// TIA Portal V19 export
FUNCTION_BLOCK "SKIDS"   // FB18, LAD
{ S7_Optimized_Access := 'TRUE' }
// stored: MemoryReserve 100, SetENOAutomatically false
   VAR
      CHILLED_SKIDS_Instance { S7_SetPoint := 'True'} : "SKIDS_LOGIC";
      START_Instance { S7_SetPoint := 'True'} : "START";
      START_Instance_COLD_SKIDS { S7_SetPoint := 'True'} : "START";
      CS_SKIDS_Instance_1 { S7_SetPoint := 'True'} : "SKIDS_LOGIC";
      START_Instance_UCH { S7_SetPoint := 'True'} : "START";
      ULTRACHILLED_SKIDS_Instance { S7_SetPoint := 'True'} : "SKIDS_LOGIC";
      ULTRACHILLED_SKIDS_Instance_1 { S7_SetPoint := 'True'} : "ULTRACHILLED_SKIDS";
      HOT_SKIDS_InstancE { S7_SetPoint := 'True'} : "SKIDS_LOGIC";
      HOT_SKIDS_Instance_1 { S7_SetPoint := 'True'} : "HOT_SKIDS";
      START_Instance_HOT_SKIDS { S7_SetPoint := 'True'} : "START";
   END_VAR
BEGIN

REGION Network 1: CHILLED SKIDS START
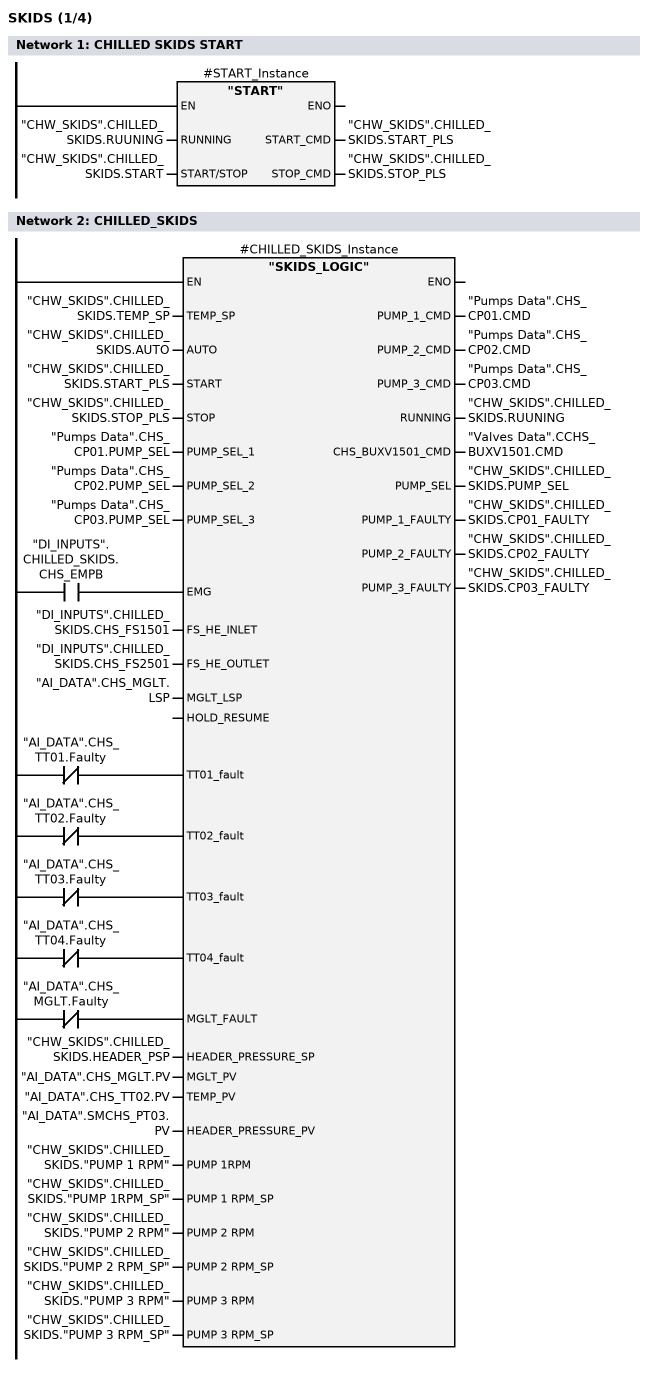
   RUNG wire#powerrail
      #START_Instance(RUNNING := "CHW_SKIDS".CHILLED_SKIDS.RUUNING, "START/STOP" := "CHW_SKIDS".CHILLED_SKIDS.START, START_CMD => "CHW_SKIDS".CHILLED_SKIDS.START_PLS, STOP_CMD => "CHW_SKIDS".CHILLED_SKIDS.STOP_PLS)
   END_RUNG
   // the same network as SCL:
   #START_Instance(RUNNING := "CHW_SKIDS".CHILLED_SKIDS.RUUNING,   // "START"
                   "START/STOP" := "CHW_SKIDS".CHILLED_SKIDS.START,
                   START_CMD => "CHW_SKIDS".CHILLED_SKIDS.START_PLS,
                   STOP_CMD => "CHW_SKIDS".CHILLED_SKIDS.STOP_PLS);
END_REGION

REGION Network 2: CHILLED_SKIDS
   RUNG wire#powerrail
      #CHILLED_SKIDS_Instance(EMG := wire#w1, TT01_fault := wire#w2, TT02_fault := wire#w3, TT03_fault := wire#w4, TT04_fault := wire#w5, MGLT_FAULT := wire#w6, TEMP_SP := "CHW_SKIDS".CHILLED_SKIDS.TEMP_SP, AUTO := "CHW_SKIDS".CHILLED_SKIDS.AUTO, START := "CHW_SKIDS".CHILLED_SKIDS.START_PLS, STOP := "CHW_SKIDS".CHILLED_SKIDS.STOP_PLS, PUMP_SEL_1 := "Pumps Data".CHS_CP01.PUMP_SEL, PUMP_SEL_2 := "Pumps Data".CHS_CP02.PUMP_SEL, PUMP_SEL_3 := "Pumps Data".CHS_CP03.PUMP_SEL, FS_HE_INLET := "DI_INPUTS".CHILLED_SKIDS.CHS_FS1501, FS_HE_OUTLET := "DI_INPUTS".CHILLED_SKIDS.CHS_FS2501, MGLT_LSP := "AI_DATA".CHS_MGLT.LSP, HOLD_RESUME :=, HEADER_PRESSURE_SP := "CHW_SKIDS".CHILLED_SKIDS.HEADER_PSP, MGLT_PV := "AI_DATA".CHS_MGLT.PV, TEMP_PV := "AI_DATA".CHS_TT02.PV, HEADER_PRESSURE_PV := "AI_DATA".SMCHS_PT03.PV, "PUMP 1RPM" := "CHW_SKIDS".CHILLED_SKIDS."PUMP 1 RPM", "PUMP 1 RPM_SP" := "CHW_SKIDS".CHILLED_SKIDS."PUMP 1RPM_SP", "PUMP 2 RPM" := "CHW_SKIDS".CHILLED_SKIDS."PUMP 2 RPM", "PUMP 2 RPM_SP" := "CHW_SKIDS".CHILLED_SKIDS."PUMP 2 RPM_SP", "PUMP 3 RPM" := "CHW_SKIDS".CHILLED_SKIDS."PUMP 3 RPM", "PUMP 3 RPM_SP" := "CHW_SKIDS".CHILLED_SKIDS."PUMP 3 RPM_SP", PUMP_1_CMD => "Pumps Data".CHS_CP01.CMD, PUMP_2_CMD => "Pumps Data".CHS_CP02.CMD, PUMP_3_CMD => "Pumps Data".CHS_CP03.CMD, RUNNING => "CHW_SKIDS".CHILLED_SKIDS.RUUNING, CHS_BUXV1501_CMD => "Valves Data".CCHS_BUXV1501.CMD, PUMP_SEL => "CHW_SKIDS".CHILLED_SKIDS.PUMP_SEL, PUMP_1_FAULTY => "CHW_SKIDS".CHILLED_SKIDS.CP01_FAULTY, PUMP_2_FAULTY => "CHW_SKIDS".CHILLED_SKIDS.CP02_FAULTY, PUMP_3_FAULTY => "CHW_SKIDS".CHILLED_SKIDS.CP03_FAULTY)
   END_RUNG
   RUNG wire#powerrail
      Contact( "DI_INPUTS".CHILLED_SKIDS.CHS_EMPB )
   END_RUNG wire#w1
   RUNG wire#powerrail
      I_Contact( "AI_DATA".CHS_TT01.Faulty )
   END_RUNG wire#w2
   RUNG wire#powerrail
      I_Contact( "AI_DATA".CHS_TT02.Faulty )
   END_RUNG wire#w3
   RUNG wire#powerrail
      I_Contact( "AI_DATA".CHS_TT03.Faulty )
   END_RUNG wire#w4
   RUNG wire#powerrail
      I_Contact( "AI_DATA".CHS_TT04.Faulty )
   END_RUNG wire#w5
   RUNG wire#powerrail
      I_Contact( "AI_DATA".CHS_MGLT.Faulty )
   END_RUNG wire#w6
   // the same network as SCL:
   #CHILLED_SKIDS_Instance(TEMP_SP := "CHW_SKIDS".CHILLED_SKIDS.TEMP_SP,   // "SKIDS_LOGIC"
                           AUTO := "CHW_SKIDS".CHILLED_SKIDS.AUTO,
                           START := "CHW_SKIDS".CHILLED_SKIDS.START_PLS,
                           STOP := "CHW_SKIDS".CHILLED_SKIDS.STOP_PLS,
                           PUMP_SEL_1 := "Pumps Data".CHS_CP01.PUMP_SEL,
                           PUMP_SEL_2 := "Pumps Data".CHS_CP02.PUMP_SEL,
                           PUMP_SEL_3 := "Pumps Data".CHS_CP03.PUMP_SEL,
                           EMG := "DI_INPUTS".CHILLED_SKIDS.CHS_EMPB,
                           FS_HE_INLET := "DI_INPUTS".CHILLED_SKIDS.CHS_FS1501,
                           FS_HE_OUTLET := "DI_INPUTS".CHILLED_SKIDS.CHS_FS2501,
                           MGLT_LSP := "AI_DATA".CHS_MGLT.LSP,
                           TT01_fault := NOT "AI_DATA".CHS_TT01.Faulty,
                           TT02_fault := NOT "AI_DATA".CHS_TT02.Faulty,
                           TT03_fault := NOT "AI_DATA".CHS_TT03.Faulty,
                           TT04_fault := NOT "AI_DATA".CHS_TT04.Faulty,
                           MGLT_FAULT := NOT "AI_DATA".CHS_MGLT.Faulty,
                           HEADER_PRESSURE_SP := "CHW_SKIDS".CHILLED_SKIDS.HEADER_PSP,
                           MGLT_PV := "AI_DATA".CHS_MGLT.PV,
                           TEMP_PV := "AI_DATA".CHS_TT02.PV,
                           HEADER_PRESSURE_PV := "AI_DATA".SMCHS_PT03.PV,
                           "PUMP 1RPM" := "CHW_SKIDS".CHILLED_SKIDS."PUMP 1 RPM",
                           "PUMP 1 RPM_SP" := "CHW_SKIDS".CHILLED_SKIDS."PUMP 1RPM_SP",
                           "PUMP 2 RPM" := "CHW_SKIDS".CHILLED_SKIDS."PUMP 2 RPM",
                           "PUMP 2 RPM_SP" := "CHW_SKIDS".CHILLED_SKIDS."PUMP 2 RPM_SP",
                           "PUMP 3 RPM" := "CHW_SKIDS".CHILLED_SKIDS."PUMP 3 RPM",
                           "PUMP 3 RPM_SP" := "CHW_SKIDS".CHILLED_SKIDS."PUMP 3 RPM_SP",
                           PUMP_1_CMD => "Pumps Data".CHS_CP01.CMD,
                           PUMP_2_CMD => "Pumps Data".CHS_CP02.CMD,
                           PUMP_3_CMD => "Pumps Data".CHS_CP03.CMD,
                           RUNNING => "CHW_SKIDS".CHILLED_SKIDS.RUUNING,
                           CHS_BUXV1501_CMD => "Valves Data".CCHS_BUXV1501.CMD,
                           PUMP_SEL => "CHW_SKIDS".CHILLED_SKIDS.PUMP_SEL,
                           PUMP_1_FAULTY => "CHW_SKIDS".CHILLED_SKIDS.CP01_FAULTY,
                           PUMP_2_FAULTY => "CHW_SKIDS".CHILLED_SKIDS.CP02_FAULTY,
                           PUMP_3_FAULTY => "CHW_SKIDS".CHILLED_SKIDS.CP03_FAULTY);
END_REGION

REGION Network 3: COLD SKIDS START
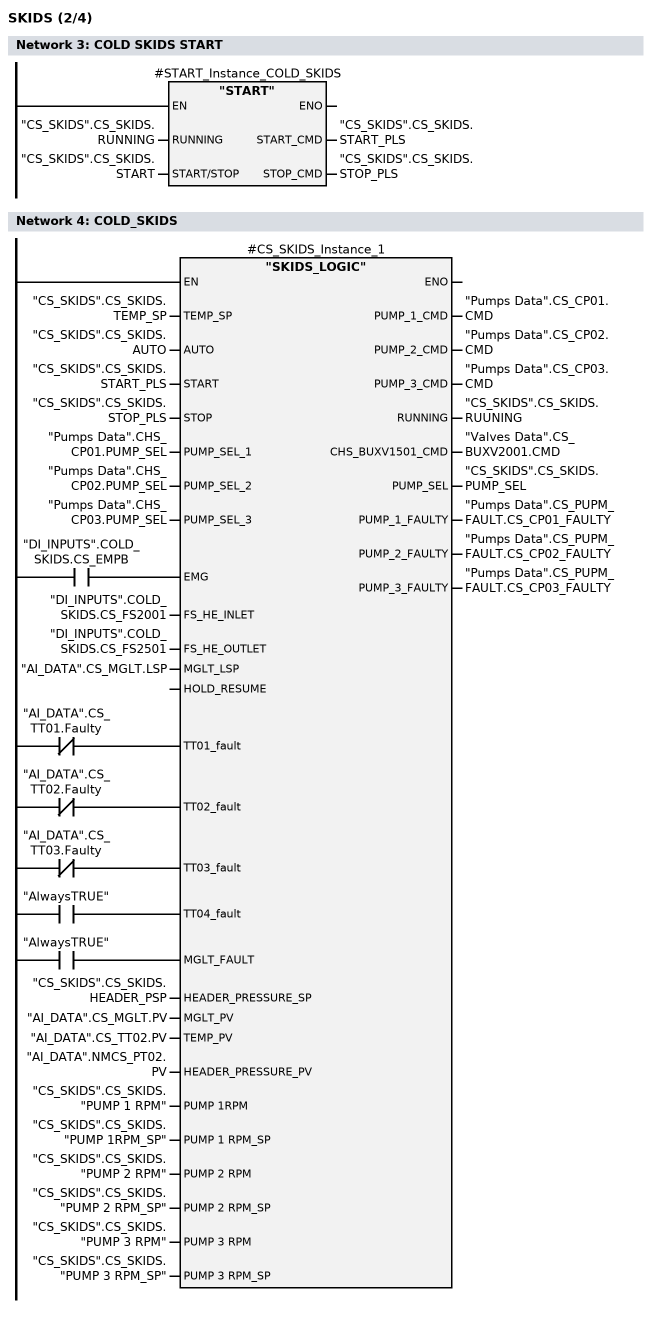
   RUNG wire#powerrail
      #START_Instance_COLD_SKIDS(RUNNING := "CS_SKIDS".CS_SKIDS.RUNNING, "START/STOP" := "CS_SKIDS".CS_SKIDS.START, START_CMD => "CS_SKIDS".CS_SKIDS.START_PLS, STOP_CMD => "CS_SKIDS".CS_SKIDS.STOP_PLS)
   END_RUNG
   // the same network as SCL:
   #START_Instance_COLD_SKIDS(RUNNING := "CS_SKIDS".CS_SKIDS.RUNNING,   // "START"
                           "START/STOP" := "CS_SKIDS".CS_SKIDS.START,
                           START_CMD => "CS_SKIDS".CS_SKIDS.START_PLS,
                           STOP_CMD => "CS_SKIDS".CS_SKIDS.STOP_PLS);
END_REGION

REGION Network 4: COLD_SKIDS
   RUNG wire#powerrail
      #CS_SKIDS_Instance_1(EMG := wire#w1, TT01_fault := wire#w2, TT02_fault := wire#w3, TT03_fault := wire#w4, TT04_fault := wire#w5, MGLT_FAULT := wire#w6, TEMP_SP := "CS_SKIDS".CS_SKIDS.TEMP_SP, AUTO := "CS_SKIDS".CS_SKIDS.AUTO, START := "CS_SKIDS".CS_SKIDS.START_PLS, STOP := "CS_SKIDS".CS_SKIDS.STOP_PLS, PUMP_SEL_1 := "Pumps Data".CHS_CP01.PUMP_SEL, PUMP_SEL_2 := "Pumps Data".CHS_CP02.PUMP_SEL, PUMP_SEL_3 := "Pumps Data".CHS_CP03.PUMP_SEL, FS_HE_INLET := "DI_INPUTS".COLD_SKIDS.CS_FS2001, FS_HE_OUTLET := "DI_INPUTS".COLD_SKIDS.CS_FS2501, MGLT_LSP := "AI_DATA".CS_MGLT.LSP, HOLD_RESUME :=, HEADER_PRESSURE_SP := "CS_SKIDS".CS_SKIDS.HEADER_PSP, MGLT_PV := "AI_DATA".CS_MGLT.PV, TEMP_PV := "AI_DATA".CS_TT02.PV, HEADER_PRESSURE_PV := "AI_DATA".NMCS_PT02.PV, "PUMP 1RPM" := "CS_SKIDS".CS_SKIDS."PUMP 1 RPM", "PUMP 1 RPM_SP" := "CS_SKIDS".CS_SKIDS."PUMP 1RPM_SP", "PUMP 2 RPM" := "CS_SKIDS".CS_SKIDS."PUMP 2 RPM", "PUMP 2 RPM_SP" := "CS_SKIDS".CS_SKIDS."PUMP 2 RPM_SP", "PUMP 3 RPM" := "CS_SKIDS".CS_SKIDS."PUMP 3 RPM", "PUMP 3 RPM_SP" := "CS_SKIDS".CS_SKIDS."PUMP 3 RPM_SP", PUMP_1_CMD => "Pumps Data".CS_CP01.CMD, PUMP_2_CMD => "Pumps Data".CS_CP02.CMD, PUMP_3_CMD => "Pumps Data".CS_CP03.CMD, RUNNING => "CS_SKIDS".CS_SKIDS.RUUNING, CHS_BUXV1501_CMD => "Valves Data".CS_BUXV2001.CMD, PUMP_SEL => "CS_SKIDS".CS_SKIDS.PUMP_SEL, PUMP_1_FAULTY => "Pumps Data".CS_PUPM_FAULT.CS_CP01_FAULTY, PUMP_2_FAULTY => "Pumps Data".CS_PUPM_FAULT.CS_CP02_FAULTY, PUMP_3_FAULTY => "Pumps Data".CS_PUPM_FAULT.CS_CP03_FAULTY)
   END_RUNG
   RUNG wire#powerrail
      Contact( "DI_INPUTS".COLD_SKIDS.CS_EMPB )
   END_RUNG wire#w1
   RUNG wire#powerrail
      I_Contact( "AI_DATA".CS_TT01.Faulty )
   END_RUNG wire#w2
   RUNG wire#powerrail
      I_Contact( "AI_DATA".CS_TT02.Faulty )
   END_RUNG wire#w3
   RUNG wire#powerrail
      I_Contact( "AI_DATA".CS_TT03.Faulty )
   END_RUNG wire#w4
   RUNG wire#powerrail
      Contact( "AlwaysTRUE" )
   END_RUNG wire#w5
   RUNG wire#powerrail
      Contact( "AlwaysTRUE" )
   END_RUNG wire#w6
   // the same network as SCL:
   #CS_SKIDS_Instance_1(TEMP_SP := "CS_SKIDS".CS_SKIDS.TEMP_SP,   // "SKIDS_LOGIC"
                        AUTO := "CS_SKIDS".CS_SKIDS.AUTO,
                        START := "CS_SKIDS".CS_SKIDS.START_PLS,
                        STOP := "CS_SKIDS".CS_SKIDS.STOP_PLS,
                        PUMP_SEL_1 := "Pumps Data".CHS_CP01.PUMP_SEL,
                        PUMP_SEL_2 := "Pumps Data".CHS_CP02.PUMP_SEL,
                        PUMP_SEL_3 := "Pumps Data".CHS_CP03.PUMP_SEL,
                        EMG := "DI_INPUTS".COLD_SKIDS.CS_EMPB,
                        FS_HE_INLET := "DI_INPUTS".COLD_SKIDS.CS_FS2001,
                        FS_HE_OUTLET := "DI_INPUTS".COLD_SKIDS.CS_FS2501,
                        MGLT_LSP := "AI_DATA".CS_MGLT.LSP,
                        TT01_fault := NOT "AI_DATA".CS_TT01.Faulty,
                        TT02_fault := NOT "AI_DATA".CS_TT02.Faulty,
                        TT03_fault := NOT "AI_DATA".CS_TT03.Faulty,
                        TT04_fault := "AlwaysTRUE",
                        MGLT_FAULT := "AlwaysTRUE",
                        HEADER_PRESSURE_SP := "CS_SKIDS".CS_SKIDS.HEADER_PSP,
                        MGLT_PV := "AI_DATA".CS_MGLT.PV,
                        TEMP_PV := "AI_DATA".CS_TT02.PV,
                        HEADER_PRESSURE_PV := "AI_DATA".NMCS_PT02.PV,
                        "PUMP 1RPM" := "CS_SKIDS".CS_SKIDS."PUMP 1 RPM",
                        "PUMP 1 RPM_SP" := "CS_SKIDS".CS_SKIDS."PUMP 1RPM_SP",
                        "PUMP 2 RPM" := "CS_SKIDS".CS_SKIDS."PUMP 2 RPM",
                        "PUMP 2 RPM_SP" := "CS_SKIDS".CS_SKIDS."PUMP 2 RPM_SP",
                        "PUMP 3 RPM" := "CS_SKIDS".CS_SKIDS."PUMP 3 RPM",
                        "PUMP 3 RPM_SP" := "CS_SKIDS".CS_SKIDS."PUMP 3 RPM_SP",
                        PUMP_1_CMD => "Pumps Data".CS_CP01.CMD,
                        PUMP_2_CMD => "Pumps Data".CS_CP02.CMD,
                        PUMP_3_CMD => "Pumps Data".CS_CP03.CMD,
                        RUNNING => "CS_SKIDS".CS_SKIDS.RUUNING,
                        CHS_BUXV1501_CMD => "Valves Data".CS_BUXV2001.CMD,
                        PUMP_SEL => "CS_SKIDS".CS_SKIDS.PUMP_SEL,
                        PUMP_1_FAULTY => "Pumps Data".CS_PUPM_FAULT.CS_CP01_FAULTY,
                        PUMP_2_FAULTY => "Pumps Data".CS_PUPM_FAULT.CS_CP02_FAULTY,
                        PUMP_3_FAULTY => "Pumps Data".CS_PUPM_FAULT.CS_CP03_FAULTY);
END_REGION

REGION Network 5: ULTRACHILLED SKIDS START
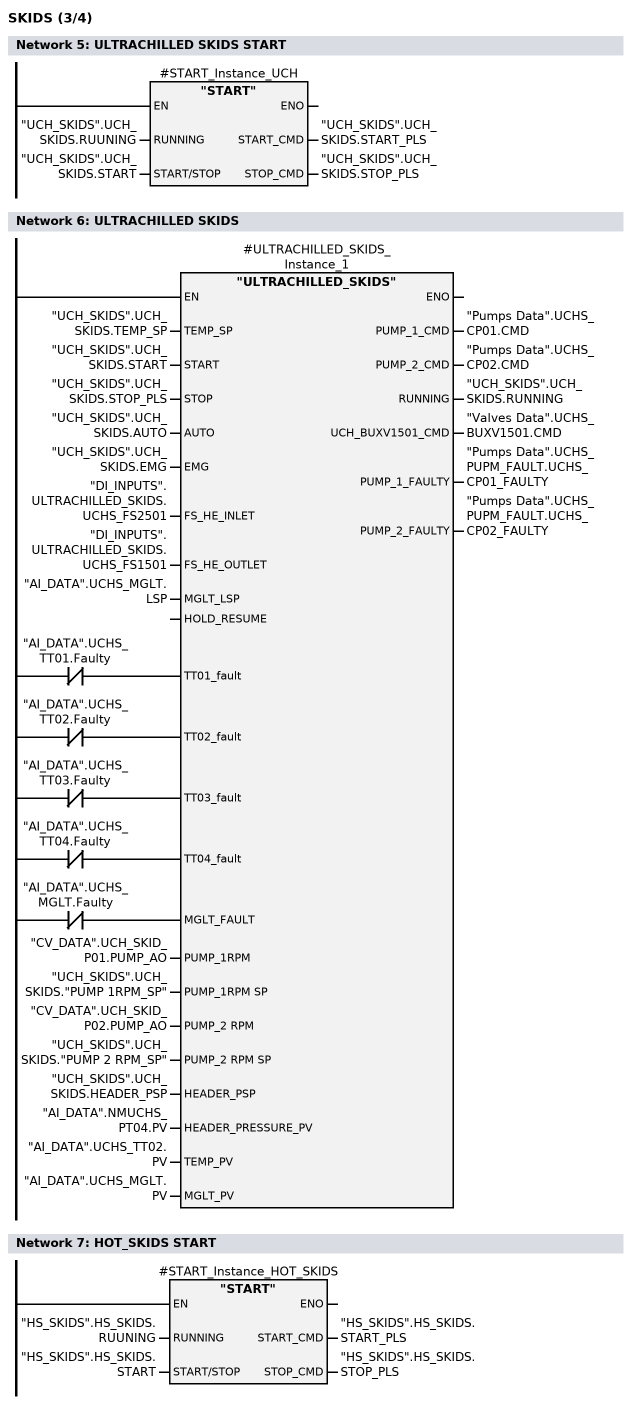
   RUNG wire#powerrail
      #START_Instance_UCH(RUNNING := "UCH_SKIDS".UCH_SKIDS.RUUNING, "START/STOP" := "UCH_SKIDS".UCH_SKIDS.START, START_CMD => "UCH_SKIDS".UCH_SKIDS.START_PLS, STOP_CMD => "UCH_SKIDS".UCH_SKIDS.STOP_PLS)
   END_RUNG
   // the same network as SCL:
   #START_Instance_UCH(RUNNING := "UCH_SKIDS".UCH_SKIDS.RUUNING,   // "START"
                       "START/STOP" := "UCH_SKIDS".UCH_SKIDS.START,
                       START_CMD => "UCH_SKIDS".UCH_SKIDS.START_PLS,
                       STOP_CMD => "UCH_SKIDS".UCH_SKIDS.STOP_PLS);
END_REGION

REGION Network 6: ULTRACHILLED SKIDS
   RUNG wire#powerrail
      #ULTRACHILLED_SKIDS_Instance_1(TT01_fault := wire#w1, TT02_fault := wire#w2, TT03_fault := wire#w3, TT04_fault := wire#w4, MGLT_FAULT := wire#w5, TEMP_SP := "UCH_SKIDS".UCH_SKIDS.TEMP_SP, START := "UCH_SKIDS".UCH_SKIDS.START, STOP := "UCH_SKIDS".UCH_SKIDS.STOP_PLS, AUTO := "UCH_SKIDS".UCH_SKIDS.AUTO, EMG := "UCH_SKIDS".UCH_SKIDS.EMG, FS_HE_INLET := "DI_INPUTS".ULTRACHILLED_SKIDS.UCHS_FS2501, FS_HE_OUTLET := "DI_INPUTS".ULTRACHILLED_SKIDS.UCHS_FS1501, MGLT_LSP := "AI_DATA".UCHS_MGLT.LSP, HOLD_RESUME :=, PUMP_1RPM := "CV_DATA".UCH_SKID_P01.PUMP_AO, "PUMP_1RPM SP" := "UCH_SKIDS".UCH_SKIDS."PUMP 1RPM_SP", "PUMP_2 RPM" := "CV_DATA".UCH_SKID_P02.PUMP_AO, "PUMP_2 RPM SP" := "UCH_SKIDS".UCH_SKIDS."PUMP 2 RPM_SP", HEADER_PSP := "UCH_SKIDS".UCH_SKIDS.HEADER_PSP, HEADER_PRESSURE_PV := "AI_DATA".NMUCHS_PT04.PV, TEMP_PV := "AI_DATA".UCHS_TT02.PV, MGLT_PV := "AI_DATA".UCHS_MGLT.PV, PUMP_1_CMD => "Pumps Data".UCHS_CP01.CMD, PUMP_2_CMD => "Pumps Data".UCHS_CP02.CMD, RUNNING => "UCH_SKIDS".UCH_SKIDS.RUNNING, UCH_BUXV1501_CMD => "Valves Data".UCHS_BUXV1501.CMD, PUMP_1_FAULTY => "Pumps Data".UCHS_PUPM_FAULT.UCHS_CP01_FAULTY, PUMP_2_FAULTY => "Pumps Data".UCHS_PUPM_FAULT.UCHS_CP02_FAULTY)
   END_RUNG
   RUNG wire#powerrail
      I_Contact( "AI_DATA".UCHS_TT01.Faulty )
   END_RUNG wire#w1
   RUNG wire#powerrail
      I_Contact( "AI_DATA".UCHS_TT02.Faulty )
   END_RUNG wire#w2
   RUNG wire#powerrail
      I_Contact( "AI_DATA".UCHS_TT03.Faulty )
   END_RUNG wire#w3
   RUNG wire#powerrail
      I_Contact( "AI_DATA".UCHS_TT04.Faulty )
   END_RUNG wire#w4
   RUNG wire#powerrail
      I_Contact( "AI_DATA".UCHS_MGLT.Faulty )
   END_RUNG wire#w5
   // the same network as SCL:
   #ULTRACHILLED_SKIDS_Instance_1(TEMP_SP := "UCH_SKIDS".UCH_SKIDS.TEMP_SP,   // "ULTRACHILLED_SKIDS"
                           START := "UCH_SKIDS".UCH_SKIDS.START,
                           STOP := "UCH_SKIDS".UCH_SKIDS.STOP_PLS,
                           AUTO := "UCH_SKIDS".UCH_SKIDS.AUTO,
                           EMG := "UCH_SKIDS".UCH_SKIDS.EMG,
                           FS_HE_INLET := "DI_INPUTS".ULTRACHILLED_SKIDS.UCHS_FS2501,
                           FS_HE_OUTLET := "DI_INPUTS".ULTRACHILLED_SKIDS.UCHS_FS1501,
                           MGLT_LSP := "AI_DATA".UCHS_MGLT.LSP,
                           TT01_fault := NOT "AI_DATA".UCHS_TT01.Faulty,
                           TT02_fault := NOT "AI_DATA".UCHS_TT02.Faulty,
                           TT03_fault := NOT "AI_DATA".UCHS_TT03.Faulty,
                           TT04_fault := NOT "AI_DATA".UCHS_TT04.Faulty,
                           MGLT_FAULT := NOT "AI_DATA".UCHS_MGLT.Faulty,
                           PUMP_1RPM := "CV_DATA".UCH_SKID_P01.PUMP_AO,
                           "PUMP_1RPM SP" := "UCH_SKIDS".UCH_SKIDS."PUMP 1RPM_SP",
                           "PUMP_2 RPM" := "CV_DATA".UCH_SKID_P02.PUMP_AO,
                           "PUMP_2 RPM SP" := "UCH_SKIDS".UCH_SKIDS."PUMP 2 RPM_SP",
                           HEADER_PSP := "UCH_SKIDS".UCH_SKIDS.HEADER_PSP,
                           HEADER_PRESSURE_PV := "AI_DATA".NMUCHS_PT04.PV,
                           TEMP_PV := "AI_DATA".UCHS_TT02.PV,
                           MGLT_PV := "AI_DATA".UCHS_MGLT.PV,
                           PUMP_1_CMD => "Pumps Data".UCHS_CP01.CMD,
                           PUMP_2_CMD => "Pumps Data".UCHS_CP02.CMD,
                           RUNNING => "UCH_SKIDS".UCH_SKIDS.RUNNING,
                           UCH_BUXV1501_CMD => "Valves Data".UCHS_BUXV1501.CMD,
                           PUMP_1_FAULTY => "Pumps Data".UCHS_PUPM_FAULT.UCHS_CP01_FAULTY,
                           PUMP_2_FAULTY => "Pumps Data".UCHS_PUPM_FAULT.UCHS_CP02_FAULTY);
END_REGION

REGION Network 7: HOT_SKIDS START
   RUNG wire#powerrail
      #START_Instance_HOT_SKIDS(RUNNING := "HS_SKIDS".HS_SKIDS.RUUNING, "START/STOP" := "HS_SKIDS".HS_SKIDS.START, START_CMD => "HS_SKIDS".HS_SKIDS.START_PLS, STOP_CMD => "HS_SKIDS".HS_SKIDS.STOP_PLS)
   END_RUNG
   // the same network as SCL:
   #START_Instance_HOT_SKIDS(RUNNING := "HS_SKIDS".HS_SKIDS.RUUNING,   // "START"
                           "START/STOP" := "HS_SKIDS".HS_SKIDS.START,
                           START_CMD => "HS_SKIDS".HS_SKIDS.START_PLS,
                           STOP_CMD => "HS_SKIDS".HS_SKIDS.STOP_PLS);
END_REGION

REGION Network 8: HOT_SKIDS
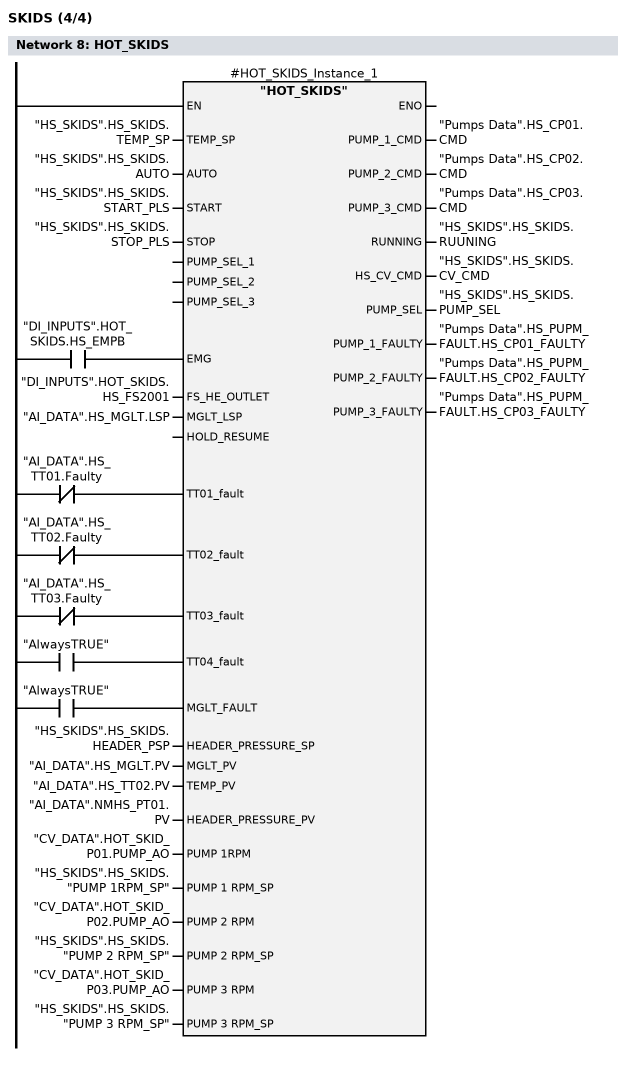
   RUNG wire#powerrail
      #HOT_SKIDS_Instance_1(EMG := wire#w1, TT01_fault := wire#w2, TT02_fault := wire#w3, TT03_fault := wire#w4, TT04_fault := wire#w5, MGLT_FAULT := wire#w6, TEMP_SP := "HS_SKIDS".HS_SKIDS.TEMP_SP, AUTO := "HS_SKIDS".HS_SKIDS.AUTO, START := "HS_SKIDS".HS_SKIDS.START_PLS, STOP := "HS_SKIDS".HS_SKIDS.STOP_PLS, PUMP_SEL_1 :=, PUMP_SEL_2 :=, PUMP_SEL_3 :=, FS_HE_OUTLET := "DI_INPUTS".HOT_SKIDS.HS_FS2001, MGLT_LSP := "AI_DATA".HS_MGLT.LSP, HOLD_RESUME :=, HEADER_PRESSURE_SP := "HS_SKIDS".HS_SKIDS.HEADER_PSP, MGLT_PV := "AI_DATA".HS_MGLT.PV, TEMP_PV := "AI_DATA".HS_TT02.PV, HEADER_PRESSURE_PV := "AI_DATA".NMHS_PT01.PV, "PUMP 1RPM" := "CV_DATA".HOT_SKID_P01.PUMP_AO, "PUMP 1 RPM_SP" := "HS_SKIDS".HS_SKIDS."PUMP 1RPM_SP", "PUMP 2 RPM" := "CV_DATA".HOT_SKID_P02.PUMP_AO, "PUMP 2 RPM_SP" := "HS_SKIDS".HS_SKIDS."PUMP 2 RPM_SP", "PUMP 3 RPM" := "CV_DATA".HOT_SKID_P03.PUMP_AO, "PUMP 3 RPM_SP" := "HS_SKIDS".HS_SKIDS."PUMP 3 RPM_SP", PUMP_1_CMD => "Pumps Data".HS_CP01.CMD, PUMP_2_CMD => "Pumps Data".HS_CP02.CMD, PUMP_3_CMD => "Pumps Data".HS_CP03.CMD, RUNNING => "HS_SKIDS".HS_SKIDS.RUUNING, HS_CV_CMD => "HS_SKIDS".HS_SKIDS.CV_CMD, PUMP_SEL => "HS_SKIDS".HS_SKIDS.PUMP_SEL, PUMP_1_FAULTY => "Pumps Data".HS_PUPM_FAULT.HS_CP01_FAULTY, PUMP_2_FAULTY => "Pumps Data".HS_PUPM_FAULT.HS_CP02_FAULTY, PUMP_3_FAULTY => "Pumps Data".HS_PUPM_FAULT.HS_CP03_FAULTY)
   END_RUNG
   RUNG wire#powerrail
      Contact( "DI_INPUTS".HOT_SKIDS.HS_EMPB )
   END_RUNG wire#w1
   RUNG wire#powerrail
      I_Contact( "AI_DATA".HS_TT01.Faulty )
   END_RUNG wire#w2
   RUNG wire#powerrail
      I_Contact( "AI_DATA".HS_TT02.Faulty )
   END_RUNG wire#w3
   RUNG wire#powerrail
      I_Contact( "AI_DATA".HS_TT03.Faulty )
   END_RUNG wire#w4
   RUNG wire#powerrail
      Contact( "AlwaysTRUE" )
   END_RUNG wire#w5
   RUNG wire#powerrail
      Contact( "AlwaysTRUE" )
   END_RUNG wire#w6
   // the same network as SCL:
   #HOT_SKIDS_Instance_1(TEMP_SP := "HS_SKIDS".HS_SKIDS.TEMP_SP,   // "HOT_SKIDS"
                         AUTO := "HS_SKIDS".HS_SKIDS.AUTO,
                         START := "HS_SKIDS".HS_SKIDS.START_PLS,
                         STOP := "HS_SKIDS".HS_SKIDS.STOP_PLS,
                         EMG := "DI_INPUTS".HOT_SKIDS.HS_EMPB,
                         FS_HE_OUTLET := "DI_INPUTS".HOT_SKIDS.HS_FS2001,
                         MGLT_LSP := "AI_DATA".HS_MGLT.LSP,
                         TT01_fault := NOT "AI_DATA".HS_TT01.Faulty,
                         TT02_fault := NOT "AI_DATA".HS_TT02.Faulty,
                         TT03_fault := NOT "AI_DATA".HS_TT03.Faulty,
                         TT04_fault := "AlwaysTRUE",
                         MGLT_FAULT := "AlwaysTRUE",
                         HEADER_PRESSURE_SP := "HS_SKIDS".HS_SKIDS.HEADER_PSP,
                         MGLT_PV := "AI_DATA".HS_MGLT.PV,
                         TEMP_PV := "AI_DATA".HS_TT02.PV,
                         HEADER_PRESSURE_PV := "AI_DATA".NMHS_PT01.PV,
                         "PUMP 1RPM" := "CV_DATA".HOT_SKID_P01.PUMP_AO,
                         "PUMP 1 RPM_SP" := "HS_SKIDS".HS_SKIDS."PUMP 1RPM_SP",
                         "PUMP 2 RPM" := "CV_DATA".HOT_SKID_P02.PUMP_AO,
                         "PUMP 2 RPM_SP" := "HS_SKIDS".HS_SKIDS."PUMP 2 RPM_SP",
                         "PUMP 3 RPM" := "CV_DATA".HOT_SKID_P03.PUMP_AO,
                         "PUMP 3 RPM_SP" := "HS_SKIDS".HS_SKIDS."PUMP 3 RPM_SP",
                         PUMP_1_CMD => "Pumps Data".HS_CP01.CMD,
                         PUMP_2_CMD => "Pumps Data".HS_CP02.CMD,
                         PUMP_3_CMD => "Pumps Data".HS_CP03.CMD,
                         RUNNING => "HS_SKIDS".HS_SKIDS.RUUNING,
                         HS_CV_CMD => "HS_SKIDS".HS_SKIDS.CV_CMD,
                         PUMP_SEL => "HS_SKIDS".HS_SKIDS.PUMP_SEL,
                         PUMP_1_FAULTY => "Pumps Data".HS_PUPM_FAULT.HS_CP01_FAULTY,
                         PUMP_2_FAULTY => "Pumps Data".HS_PUPM_FAULT.HS_CP02_FAULTY,
                         PUMP_3_FAULTY => "Pumps Data".HS_PUPM_FAULT.HS_CP03_FAULTY);
END_REGION
END_FUNCTION_BLOCK
